FUNCTION_BLOCK FTS_MCGearOut
VAR_IN_OUT
	stSlaveAxis: ST_Axis;
END_VAR
VAR_INPUT
	bExecute: BOOL;
END_VAR
VAR_OUTPUT
	bBusy: BOOL;
	bDone: BOOL;
	bError: BOOL;
	nErrorId: UDINT;
END_VAR
VAR
	_nStep: INT;
	_fbTrig: R_TRIG;
	_fbDoneTon: TON;
END_VAR
VAR CONSTANT
	tcDoneTime: TIME := TIME#100ms;
	tcWaitTime: TIME := TIME#16m40s0ms;
END_VAR

_fbTrig(CLK:=bExecute , Q=> );
IF _fbTrig.Q AND(_nStep=0)THEN
	_nStep:=10;
END_IF


CASE _nStep  OF 
	0:
	    IF NOT bExecute THEN 
		   bError:=FALSE;
		   nErrorId:=0;
		   bDone:=FALSE;
		   
	    END_IF
	    RETURN ;
		
    10:
	    
		bBusy:=TRUE;
		bDone:=FALSE;
		bError:=FALSE;
		nErrorId:=0;
		stSlaveAxis.stPLCTONC.eCommand:=E_Command.COMMAND_GEAROUT;  //03.11
		_nStep:=20;
	20:
	    bBusy:=FALSE;
	    bDone:=TRUE;
		IF NOT stSlaveAxis.stAxisStatus.bSynchronizedMotion  THEN 
		   stSlaveAxis.stPLCTONC.eCommand:=E_Command.COMMAND_IDLE;  //03.11
		END_IF
	   // _fbDoneTon(IN:=FALSE, PT:=tcDoneTime , Q=> , ET=> );
		IF bExecute  THEN 
			_nStep:=0;
		ELSE
			_nStep:=30;
		END_IF
	    
    30:
	    //_fbDoneTon(IN:=TRUE, PT:=tcDoneTime , Q=> , ET=> );
      // IF _fbDoneTon.Q THEN
		  bDone:=FALSE;
		  _fbDoneTon(IN:=FALSE, PT:=tcDoneTime , Q=> , ET=> );
		  _nStep:=0;
		  
	  // END_IF
	
	100:
	     bBusy:=FALSE;
	     bError:=TRUE;
	     stSlaveAxis.stAxisStatus.bError:=TRUE;
	     _nStep:=0;
	

END_CASE

END_FUNCTION_BLOCK

(* stored: Version 1.1.0.1, ProductVersion 3.1.4024.12
   POU FTS_MCGearOut: Id {22e0a6ad-8b6d-4d43-b2da-bc874f489751}, SpecialFunc None *)
